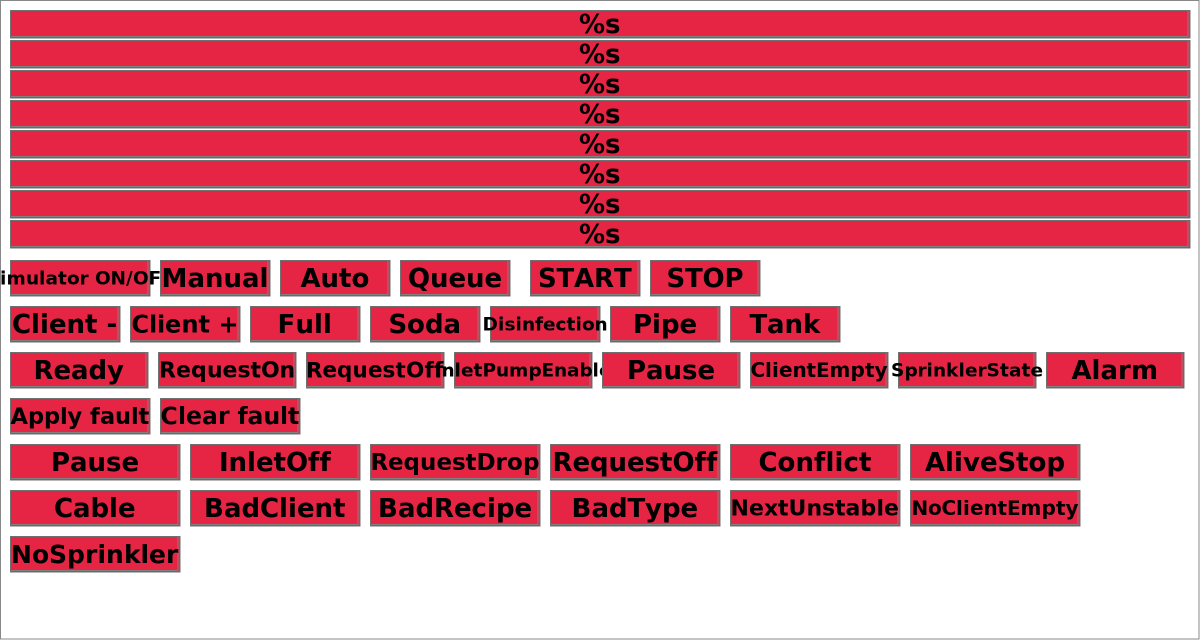
VISUALIZATION vis_SiemensSim  // 1200x640
    Button (10,10 1180x28), "%s", text variable: g_Anybus.fbSim.sSim
    Button (10,40 1180x28), "%s", text variable: g_Anybus.fbSim.sMode
    Button (10,70 1180x28), "%s", text variable: g_Anybus.fbSim.sClient
    Button (10,100 1180x28), "%s", text variable: g_Anybus.fbSim.sFault
    Button (10,130 1180x28), "%s", text variable: g_Anybus.fbSim.sFromCip
    Button (10,160 1180x28), "%s", text variable: g_Anybus.fbSim.sToCip
    Button (10,190 1180x28), "%s", text variable: g_Anybus.fbSim.sManual
    Button (10,220 1180x28), "%s", text variable: g_Anybus.fbSim.sInterface
    Button (10,260 140x36), "Simulator ON/OFF"
        OnMouseClick: execute { g_Anybus.bSimEnable:=NOT g_Anybus.bSimEnable; }
    Button (160,260 110x36), "Manual"
        OnMouseClick: execute { g_Anybus.fbSim.eMode:=E_Sim_Mode.eManual; }
    Button (280,260 110x36), "Auto"
        OnMouseClick: execute { g_Anybus.fbSim.eMode:=E_Sim_Mode.eAuto; }
    Button (400,260 110x36), "Queue"
        OnMouseClick: execute { g_Anybus.fbSim.eMode:=E_Sim_Mode.eQueue; }
    Button (530,260 110x36), "START"
        OnMouseClick: execute { g_Anybus.fbSim.bStart:=TRUE; }
    Button (650,260 110x36), "STOP"
        OnMouseClick: execute { g_Anybus.fbSim.bStop:=TRUE; }
    Button (10,306 110x36), "Client -"
        OnMouseClick: execute { IF g_Anybus.fbSim.stClient.nClient>1 THEN g_Anybus.fbSim.stClient.nClient:=g_Anybus.fbSim.stClient.nClient-1; END_IF }
    Button (130,306 110x36), "Client +"
        OnMouseClick: execute { IF g_Anybus.fbSim.stClient.nClient<30 THEN g_Anybus.fbSim.stClient.nClient:=g_Anybus.fbSim.stClient.nClient+1; END_IF }
    Button (250,306 110x36), "Full"
        OnMouseClick: execute { g_Anybus.fbSim.stClient.eRecipe:=E_Anybus_RecipeType.eFull; }
    Button (370,306 110x36), "Soda"
        OnMouseClick: execute { g_Anybus.fbSim.stClient.eRecipe:=E_Anybus_RecipeType.eDetergent; }
    Button (490,306 110x36), "Disinfection"
        OnMouseClick: execute { g_Anybus.fbSim.stClient.eRecipe:=E_Anybus_RecipeType.eDisinfectionOnly; }
    Button (610,306 110x36), "Pipe"
        OnMouseClick: execute { g_Anybus.fbSim.stClient.eType:=E_Anybus_ClientType.ePipe; }
    Button (730,306 110x36), "Tank"
        OnMouseClick: execute { g_Anybus.fbSim.stClient.eType:=E_Anybus_ClientType.eTank; }
    Button (10,352 138x36), "Ready"
        OnMouseClick: execute { g_Anybus.fbSim.stManual.bReady:=NOT g_Anybus.fbSim.stManual.bReady; }
    Button (158,352 138x36), "RequestOn"
        OnMouseClick: execute { g_Anybus.fbSim.stManual.bRequestOn:=NOT g_Anybus.fbSim.stManual.bRequestOn; }
    Button (306,352 138x36), "RequestOff"
        OnMouseClick: execute { g_Anybus.fbSim.stManual.bRequestOff:=NOT g_Anybus.fbSim.stManual.bRequestOff; }
    Button (454,352 138x36), "InletPumpEnable"
        OnMouseClick: execute { g_Anybus.fbSim.stManual.bInletPumpEnable:=NOT g_Anybus.fbSim.stManual.bInletPumpEnable; }
    Button (602,352 138x36), "Pause"
        OnMouseClick: execute { g_Anybus.fbSim.stManual.bPause:=NOT g_Anybus.fbSim.stManual.bPause; }
    Button (750,352 138x36), "ClientEmpty"
        OnMouseClick: execute { g_Anybus.fbSim.stManual.bClientEmpty:=NOT g_Anybus.fbSim.stManual.bClientEmpty; }
    Button (898,352 138x36), "SprinklerState"
        OnMouseClick: execute { g_Anybus.fbSim.stManual.bSprinklerState:=NOT g_Anybus.fbSim.stManual.bSprinklerState; }
    Button (1046,352 138x36), "Alarm"
        OnMouseClick: execute { g_Anybus.fbSim.stManual.bAlarm:=NOT g_Anybus.fbSim.stManual.bAlarm; }
    Button (10,398 140x36), "Apply fault"
        OnMouseClick: execute { g_Anybus.fbSim.bFaultOn:=TRUE; }
    Button (160,398 140x36), "Clear fault"
        OnMouseClick: execute { g_Anybus.fbSim.bFaultOn:=FALSE; }
    Button (10,444 170x36), "Pause"
        OnMouseClick: execute { g_Anybus.fbSim.eFault:=E_Sim_Fault.ePause; }
    Button (190,444 170x36), "InletOff"
        OnMouseClick: execute { g_Anybus.fbSim.eFault:=E_Sim_Fault.eInletOff; }
    Button (370,444 170x36), "RequestDrop"
        OnMouseClick: execute { g_Anybus.fbSim.eFault:=E_Sim_Fault.eRequestDrop; }
    Button (550,444 170x36), "RequestOff"
        OnMouseClick: execute { g_Anybus.fbSim.eFault:=E_Sim_Fault.eRequestOff; }
    Button (730,444 170x36), "Conflict"
        OnMouseClick: execute { g_Anybus.fbSim.eFault:=E_Sim_Fault.eConflict; }
    Button (910,444 170x36), "AliveStop"
        OnMouseClick: execute { g_Anybus.fbSim.eFault:=E_Sim_Fault.eAliveStop; }
    Button (10,490 170x36), "Cable"
        OnMouseClick: execute { g_Anybus.fbSim.eFault:=E_Sim_Fault.eCable; }
    Button (190,490 170x36), "BadClient"
        OnMouseClick: execute { g_Anybus.fbSim.eFault:=E_Sim_Fault.eBadClient; }
    Button (370,490 170x36), "BadRecipe"
        OnMouseClick: execute { g_Anybus.fbSim.eFault:=E_Sim_Fault.eBadRecipe; }
    Button (550,490 170x36), "BadType"
        OnMouseClick: execute { g_Anybus.fbSim.eFault:=E_Sim_Fault.eBadType; }
    Button (730,490 170x36), "NextUnstable"
        OnMouseClick: execute { g_Anybus.fbSim.eFault:=E_Sim_Fault.eNextUnstable; }
    Button (910,490 170x36), "NoClientEmpty"
        OnMouseClick: execute { g_Anybus.fbSim.eFault:=E_Sim_Fault.eNoClientEmpty; }
    Button (10,536 170x36), "NoSprinkler"
        OnMouseClick: execute { g_Anybus.fbSim.eFault:=E_Sim_Fault.eNoSprinkler; }
END_VISUALIZATION

// ---- 03 Project/vis_Main.TcVIS
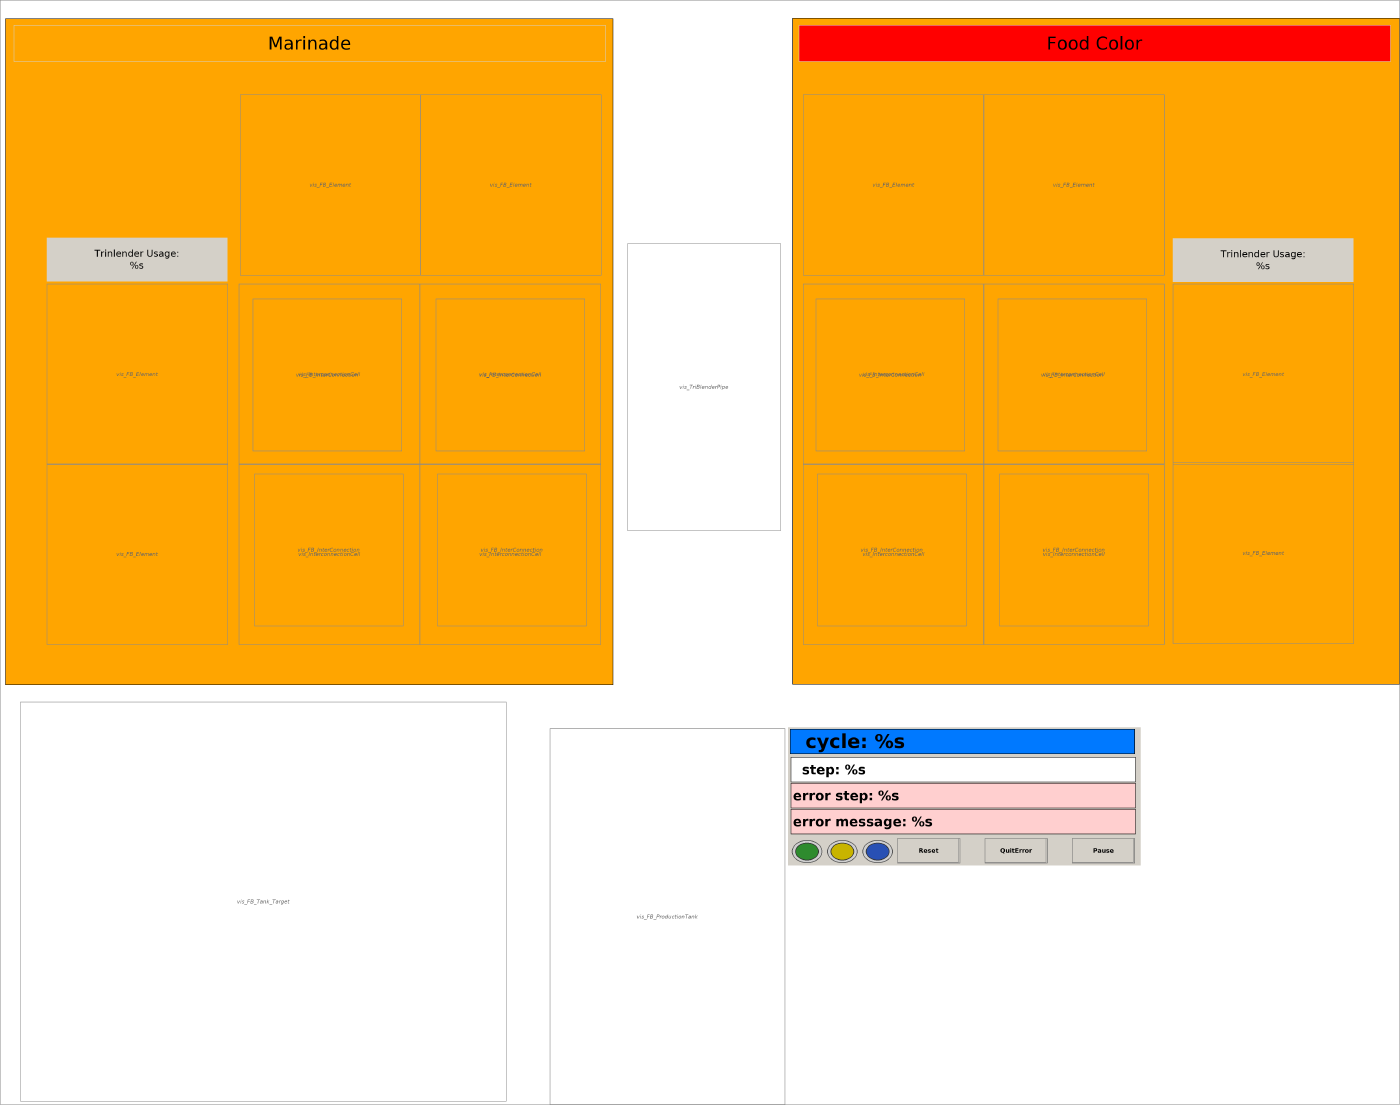
VISUALIZATION vis_Main  // 2638x2083
    Rectangle (1493,34 1145x1256)
    Frame (1513,178 341x341)
        shows vis_FB_Element(fb := fbElement[E_Element_List.eTank_3])
    Frame (1853,178 341x341)
        shows vis_FB_Element(fb := fbElement[E_Element_List.eTank_4])
    Frame (2210,535 341x341)
        shows vis_FB_Element(fb := fbElement[E_Element_List.eTriBlender_Color])
    Frame (2210,872 341x341)
        shows vis_FB_Element(fb := fbElement[E_Element_List.eLine_Color])
    Frame (1513,535 341x341)
        shows vis_InterconnectionCell()
    Frame (1853,535 341x341)
        shows vis_InterconnectionCell()
    Frame (1513,874 341x341)
        shows vis_InterconnectionCell()
    Frame (1853,874 341x341)
        shows vis_InterconnectionCell()
    Frame (1537,563 281x287)
        shows vis_FB_InterConnection(fb := fbIntCon_TriB_T3_Color)
    Frame (1880,563 281x287)
        shows vis_FB_InterConnection(fb := fbIntCon_TriB_T4_Color)
    Frame (1540,893 281x287)
        shows vis_FB_InterConnection(fb := fbIntCon_ProL_T3_Color)
    Frame (1883,893 281x287)
        shows vis_FB_InterConnection(fb := fbIntCon_ProL_T4_Color)
    Textfield (1505,47 1115x69), "Food Color"
    Group (10,35 1145x1256)
        Rectangle (0,0 1145x1256)
        Frame (442,143 341x341)
            shows vis_FB_Element(fb := fbElement[E_Element_List.eTank_1])
        Frame (782,143 341x341)
            shows vis_FB_Element(fb := fbElement[E_Element_List.eTank_2])
        Frame (78,500 341x341)
            shows vis_FB_Element(fb := fbElement[E_Element_List.eTriBlender_Marinada])
        Frame (78,839 341x341)
            shows vis_FB_Element(fb := fbElement[E_Element_List.eLine_Marinada])
        Frame (440,500 341x341)
            shows vis_InterconnectionCell()
        Frame (781,500 341x341)
            shows vis_InterconnectionCell()
        Frame (440,839 341x341)
            shows vis_InterconnectionCell()
        Frame (781,839 341x341)
            shows vis_InterconnectionCell()
        Frame (466,528 281x287)
            shows vis_FB_InterConnection(fb := fbIntCon_TriB_T1_Marin)
        Frame (811,528 281x287)
            shows vis_FB_InterConnection(fb := fbIntCon_TriB_T2_Marin)
        Frame (469,858 281x287)
            shows vis_FB_InterConnection(fb := fbIntCon_ProL_T1_Marin)
        Frame (814,858 281x287)
            shows vis_FB_InterConnection(fb := fbIntCon_ProL_T2_Marin)
        Textfield (16,12 1115x69), "Marinade"
        Textfield (78,413 340x82), "Trinlender Usage: %s", colour toggle: eTriBlenderUsage=E_TriBlenderUsage.eColor_Standby OR eTriBlenderUsage=E_TriBlenderUsage.eColor_T3 OR eTriBlenderUsage=E_TriBlenderUsage.eColor_T4, text list: 'TextList_TriBlenderUsage', text index: eTriBlenderUsage
    Textfield (2210,449 340x82), "Trinlender Usage: %s", colour toggle: eTriBlenderUsage=E_TriBlenderUsage.eMarinada_Standby OR eTriBlenderUsage=E_TriBlenderUsage.eMarinada_T1 OR eTriBlenderUsage=E_TriBlenderUsage.eMarinada_T2, text list: 'TextList_TriBlenderUsage', text index: eTriBlenderUsage
    Frame (1182,459 289x541)
        shows vis_TriBlenderPipe()
    Frame (1485,1371 664x260)
        shows vis_Cycle_Control_1(fb := fbTank1, sName := 'T1 Marinade')
    Frame (1036,1373 443x710)
        shows vis_FB_ProductionTank(fb := fbTank1)
    Frame (38,1323 916x753)
        shows vis_FB_Tank_Target(fb := fbTank1.fbTarget)
END_VISUALIZATION

// ---- GlobalTextList.TcGTLO
TEXTLIST GlobalTextList
  440 = '   message'
  1783 = '  cycle: %s'
  374 = '  step: %s'
  662 = ' %s'
  491 = '#%d'
  1694 = '%1.2f'
  153 = '%d'
  887 = '%s'
  553 = '%S'
  140 = '1/0'
  914 = '5s'
  1075 = 'Act Errors'
  1902 = 'Act State'
  690 = 'Actual'
  594 = 'Actual Errors'
  714 = 'All'
  975 = 'arCIP_RequestBufer[INDEX].eCIP_Type'
  286 = 'Auto'
  1263 = 'Axis'
  3209 = 'base time: %2.1f [sec]'
  9116 = 'ByPass'
  413 = 'bypass'
  743 = 'Cheesy Bites'
  749 = 'Cheesy Cut'
  396 = 'CIP'
  254 = 'CIP Type'
  416 = 'CIP1'
  878 = 'CIP3'
  68 = 'CIP5'
  201 = 'clean'
  677 = 'Client'
  673 = 'Close'
  1128 = 'close'
  1303 = 'Close sensor'
  8 = 'Close Sensor state'
  176 = 'Close valve'
  4398 = 'Close:'
  2046 = 'Compressor'
  520 = 'Connect'
  755 = 'Cream'
  472 = 'Crean Empty'
  742 = 'Create\nRecipe'
  1961 = 'Create Default\nRecipe'
  761 = 'Crown'
  186 = 'dealy: %.2f [sec] '
  820 = 'Default pos'
  778 = 'delay: %.2f [sec] '
  817 = 'Delete'
  713 = 'Delete\nRecipe'
  720 = 'Device 1'
  726 = 'Device 2'
  732 = 'Device 3'
  738 = 'Device 4'
  919 = 'Device Name'
  785 = 'Device State'
  178 = 'Disconnect'
  647 = 'Dissolving Done'
  47 = 'Done'
  3155 = 'Door\n#1\n'
  615 = 'Down'
  175 = 'Drain'
  460 = 'Element'
  112 = 'Emergency'
  1424 = 'Emergency Stop and Interlock'
  956 = 'EMO'
  1787 = 'Err'
  232 = 'err: %x'
  249 = 'ErrID'
  892 = 'Error'
  2981 = 'Error code: %s'
  595 = 'Error History'
  253 = 'Error Message'
  386 = 'error message: %s'
  896 = 'Error message: %s'
  5 = 'error reason: %s'
  304 = 'error step: %s'
  114 = 'Errors'
  5489 = 'Errors Search\nBuffer'
  105 = 'Errors: %d'
  3404 = 'ES Bypass'
  767 = 'Flour'
  752 = 'Food Color'
  2114 = 'Get\nLast Err'
  694 = 'History'
  756 = 'History Errors'
  3107 = 'Initialization'
  410 = 'Interlock'
  1912 = 'Interlock\nZone#1'
  4542 = 'Intilize'
  2697 = 'Last Return:'
  251 = 'Level'
  985 = 'Line'
  315 = 'link: %s'
  971 = 'Load\nRecipe'
  1122 = 'Load Recipe\nfrom file'
  135 = 'Local'
  70 = 'Main'
  2930 = 'Man'
  245 = 'Manual'
  534 = 'Marinade'
  104 = 'max: %.2f [sec] '
  11600 = 'Memo PB State'
  1148 = 'Message:'
  918 = 'min: %.2f [sec] '
  252 = 'Module Description'
  773 = 'Mozza'
  4048 = 'Mute'
  2718 = 'N'
  2076 = 'New Recipe Name:'
  920 = 'No'
  721 = 'not clean'
  181 = 'Off'
  2479 = 'OFF'
  922 = 'on'
  1164 = 'On duty: %0.1f [%]'
  952 = 'Open'
  255 = 'open'
  4392 = 'Open :'
  1663 = 'Open sensor'
  128 = 'Open Sensor state'
  197 = 'Open valve'
  779 = 'Open1'
  784 = 'Open2'
  790 = 'Open3'
  796 = 'Open4'
  444 = 'Outlet'
  1703 = 'P'
  664 = 'Password: %s'
  9135 = 'Path:'
  313 = 'Pause'
  659 = 'Pause History'
  821 = 'Piston Param'
  692 = 'piston: %s'
  704 = 'Play'
  106 = 'PLC Ver: %s'
  1953 = 'POU name: %s'
  157 = 'process: %s'
  687 = 'product'
  240 = 'Production'
  48 = 'QuitError'
  117 = 'R'
  231 = 'Ready'
  942 = 'Recipe'
  908 = 'recipe: %s'
  3336 = 'ReInit'
  2325 = 'Release ES'
  2568 = 'Reload'
  746 = 'Request Local'
  190 = 'Request Local Detergent'
  391 = 'Request Local Full'
  795 = 'request: %s'
  650 = 'Reset'
  264 = 'Reset\nErr'
  928 = 'Reset Errors'
  429 = 'Resume'
  4367 = 'Root Folder:'
  593 = 'Run'
  522 = 'Save Recipe\nto File'
  1817 = 'Save Recipe\nto file'
  1340 = 'Search'
  2084 = 'Selected Recipe:'
  2934 = 'Semi'
  1537 = 'sensor'
  183 = 'Sensor \nexist'
  814 = 'Sesame'
  953 = 'short state: %s'
  2834 = 'Standby'
  36 = 'Start Production'
  134 = 'state time: %s'
  2993 = 'state: %s'
  976 = 'status: %s'
  14674 = 'Stop\nReset All'
  812 = 'Stop Production'
  643 = 'T.C  logo '
  5392 = 'Table Index:'
  750 = 'Test'
  526 = 'Time'
  80 = 'Timing'
  1281 = 'ToBe Done'
  563 = 'TriBlender'
  96 = 'TriBlenDer'
  451 = 'Trinlender Usage:\n%s'
  915 = 'Type'
  316 = 'Up'
  745 = 'User: %s'
  810 = 'Valve'
  927 = 'Variable Name'
  936 = 'Variable Value'
  802 = 'Wet'
  808 = 'Wrap'
END_TEXTLIST
